(* PLC project fbd_seal_in, Anonymous Benchmark Suite 1.0 *)
(* stored: creationDateTime 2026-08-26T00:00:00 *)

PROGRAM drive
  VAR_INPUT
    Start : BOOL;
    Stop : BOOL;
  END_VAR
  VAR_OUTPUT
    Run : BOOL;
  END_VAR

(* FBD diagram, written out as Structured Text *)
Run := (Start OR Run) AND NOT Stop;
END_PROGRAM

CONFIGURATION Config0
  RESOURCE Res0 ON PLC
    TASK tcyclic(INTERVAL := T#10ms, PRIORITY := 0);
    PROGRAM inst0 WITH tcyclic : drive;
  END_RESOURCE
END_CONFIGURATION
